// TIA Portal V21 export
// export: Created 2026-11-18T10:00:00.0000000Z, ExportSetting None
FUNCTION_BLOCK "FB_Conveyor"   // FB10, LAD
{ S7_Optimized_Access := 'TRUE' }
// stored: MemoryReserve 100, SetENOAutomatically false
   VAR_INPUT
      Start : Bool;
      Stop : Bool;
      Direction : Bool;
      Speed : Real;
   END_VAR
   VAR_OUTPUT
      Motor : Bool;
      Fault : Bool;
   END_VAR
   VAR
      T_Startup : TON_TIME;
      Startup_Time : Time;
      Started_Up : Bool;
      Ready : Bool;
      Moving : Bool;
      Ack_P : Bool;
      Temp_High : Bool;
      Belt_Running : Bool;
   END_VAR
   VAR_TEMP   // added for the SCL form of the ladder/FBD networks
      _w1 : Bool;
      _w2 : Bool;
   END_VAR
BEGIN

REGION Network 1: Připravenost dopravníku
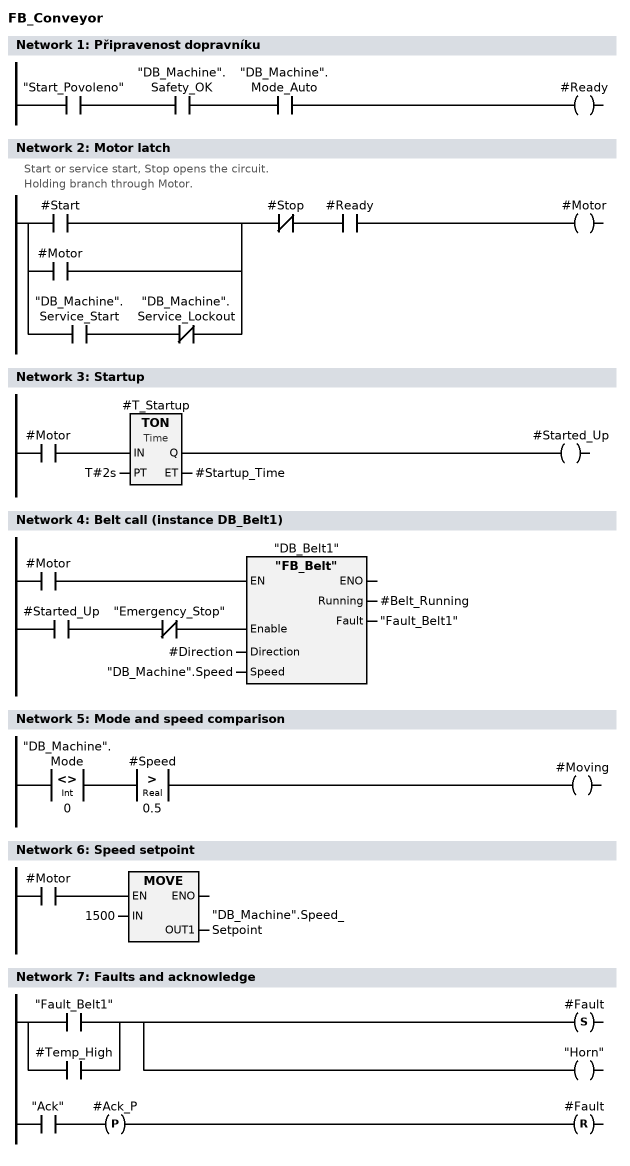
   RUNG wire#powerrail
      Contact( "Start_Povoleno" )
      Contact( "DB_Machine".Safety_OK )
      Contact( "DB_Machine".Mode_Auto )
      Coil( #Ready )
   END_RUNG
   // the same network as SCL:
   #Ready := "Start_Povoleno" AND "DB_Machine".Safety_OK AND "DB_Machine".Mode_Auto;
END_REGION

REGION Network 2: Motor latch
   // Start or service start, Stop opens the circuit.
   // Holding branch through Motor.
   #Motor := (#Start OR #Motor OR ("DB_Machine".Service_Start AND NOT "DB_Machine".Service_Lockout)) AND NOT #Stop AND #Ready;
END_REGION

REGION Network 3: Startup
   RUNG wire#powerrail
      Contact( #Motor )
      { S7_Templates := "time_type := Time" } #T_Startup.TON(pt := T#2s, et => #Startup_Time)
      Coil( #Started_Up )
   END_RUNG
   // the same network as SCL:
   #T_Startup(IN := #Motor, PT := T#2s, ET => #Startup_Time);   // TON
   #Started_Up := #T_Startup.Q;
END_REGION

REGION Network 4: Belt call (instance DB_Belt1)
   IF #Motor THEN
       "DB_Belt1"(Enable := #Started_Up AND NOT "Emergency_Stop",   // "FB_Belt"
                  Direction := #Direction,
                  Speed := "DB_Machine".Speed,
                  Running => #Belt_Running,
                  Fault => "Fault_Belt1");
   END_IF;
END_REGION

REGION Network 5: Mode and speed comparison
   RUNG wire#powerrail
      { S7_Templates := "SrcType := Int" } NE_Contact(in1 := "DB_Machine".Mode, in2 := 0)
      { S7_Templates := "SrcType := Real" } GT_Contact(in1 := #Speed, in2 := 0.5)
      Coil( #Moving )
   END_RUNG
   // the same network as SCL:
   #Moving := ("DB_Machine".Mode <> 0) AND (#Speed > 0.5);
END_REGION

REGION Network 6: Speed setpoint
   RUNG wire#powerrail
      Contact( #Motor )
      Move(in := 1500, out1 => "DB_Machine".Speed_Setpoint)
   END_RUNG
   // the same network as SCL:
   IF #Motor THEN "DB_Machine".Speed_Setpoint := 1500; END_IF;
END_REGION

REGION Network 7: Faults and acknowledge
   #_w1 := "Ack" AND NOT #Ack_P;   // rising edge
   #Ack_P := "Ack";
   IF #_w1 THEN #Fault := FALSE; END_IF;
   #_w2 := "Fault_Belt1" OR #Temp_High;
   IF #_w2 THEN #Fault := TRUE; END_IF;
   "Horn" := #_w2;
END_REGION
END_FUNCTION_BLOCK
